{attribute 'qualified_only'}
VAR_GLOBAL CONSTANT
    MODEF_SERVO_ENABLE : UINT := 16#0001;          (* bit0 *)
    MODEF_EXPERIMENT_START_REQ : UINT := 16#0002;  (* bit1 *)
    HEARTBEAT_TIMEOUT_TICKS : UDINT := 50;         (* 10 ms task * 50 = 500 ms *)

END_VAR

VAR_GLOBAL
    {attribute 'linkalways'}
    modeFlags : UINT := 0;
    resetReq : BOOL := FALSE;
    resetAckCounter : UDINT := 0;
    hostHeartbeatCounter : UDINT := 0;
    watchdogTripCounter : UDINT := 0;
    experimentActive : BOOL := FALSE;
    loggerFileReleased : BOOL := FALSE;
    loggerErrorCode : UDINT := 0;
    modeState : E_ModeState := E_ModeState.IDLE;
END_VAR

(* stored: Version 1.1.0.1
   GVL GVL_MODE: Id {4e4b78e9-90d4-4b53-9647-8f59e8f34bd4} *)
